(* IEC 61131-3 sources: TIA2AX/tests/test_projects/expected/HW_DiscoverGroups/PLC_2, 6 files *)

(* ---- HwInputs.st ---- *)
TYPE
	HwInputs : STRUCT
		PLC_2_10A_1 AT %B7 : WORD;
		PLC_2_10A_2 AT %B9 : WORD;
		PLC_2_10A_3 AT %B11 : WORD;
		PLC_2_10A_4 AT %B13 : WORD;
		PLC_2_10A_5 AT %B15 : WORD;
		PLC_2_10A_6 AT %B17 : WORD;
		_10A_16_10A_2 AT %B19 : BYTE;
		_10A_16_10A_3 AT %B20 : BYTE;
		_10A_16_10A_4 AT %B21 : BYTE;
		_10A_16_10A_5 AT %B22 : BYTE;
		_10A_16_10A_6 AT %B23 : BYTE;
		_10A_20_10A_2 AT %B24 : BYTE;
		_10A_20_10A_3 AT %B25 : BYTE;
		_10A_20_10A_4 AT %B26 : BYTE;
		_10A_20_10A_5 AT %B27 : BYTE;
		_10A_20_10A_6 AT %B28 : BYTE;
		_10A_12_10A_2 AT %B2 : BYTE;
		_10A_12_10A_3 AT %B3 : BYTE;
		_10A_12_10A_4 AT %B4 : BYTE;
		_10A_12_10A_5 AT %B5 : BYTE;
		_10A_12_10A_6 AT %B6 : BYTE;
	END_STRUCT;
END_TYPE

(* ---- HwOutputs.st ---- *)
TYPE
	HwOutputs : STRUCT
		PLC_2_10A_7 AT %B7 : WORD;
		PLC_2_10A_8 AT %B9 : WORD;
		PLC_2_10A_9 AT %B11 : WORD;
		PLC_2_10A_10 AT %B13 : WORD;
		PLC_2_10A_11 AT %B15 : WORD;
		PLC_2_10A_12 AT %B17 : WORD;
		_10A_16_10A_7 AT %B19 : BYTE;
		_10A_16_10A_8 AT %B20 : BYTE;
		_10A_16_10A_9 AT %B21 : BYTE;
		_10A_16_10A_10 AT %B22 : BYTE;
		_10A_16_10A_11 AT %B23 : BYTE;
		_10A_20_10A_7 AT %B24 : BYTE;
		_10A_20_10A_8 AT %B25 : BYTE;
		_10A_20_10A_9 AT %B26 : BYTE;
		_10A_20_10A_10 AT %B27 : BYTE;
		_10A_20_10A_11 AT %B28 : BYTE;
		_10A_12_10A_7 AT %B2 : BYTE;
		_10A_12_10A_8 AT %B3 : BYTE;
		_10A_12_10A_9 AT %B4 : BYTE;
		_10A_12_10A_10 AT %B5 : BYTE;
		_10A_12_10A_11 AT %B6 : BYTE;
	END_STRUCT;
END_TYPE

(* ---- PlcInputs.st ---- *)
TYPE
	PlcInputs : STRUCT
		PLC_2_10A_1 : WORD;
		PLC_2_10A_2 : WORD;
		PLC_2_10A_3 : WORD;
		PLC_2_10A_4 : WORD;
		PLC_2_10A_5 : WORD;
		PLC_2_10A_6 : WORD;
		_10A_16_10A_2 : BYTE;
		_10A_16_10A_3 : BYTE;
		_10A_16_10A_4 : BYTE;
		_10A_16_10A_5 : BYTE;
		_10A_16_10A_6 : BYTE;
		_10A_20_10A_2 : BYTE;
		_10A_20_10A_3 : BYTE;
		_10A_20_10A_4 : BYTE;
		_10A_20_10A_5 : BYTE;
		_10A_20_10A_6 : BYTE;
		_10A_12_10A_2 : BYTE;
		_10A_12_10A_3 : BYTE;
		_10A_12_10A_4 : BYTE;
		_10A_12_10A_5 : BYTE;
		_10A_12_10A_6 : BYTE;
	END_STRUCT;
END_TYPE

(* ---- PlcOutputs.st ---- *)
TYPE
	PlcOutputs : STRUCT
		PLC_2_10A_7 : WORD;
		PLC_2_10A_8 : WORD;
		PLC_2_10A_9 : WORD;
		PLC_2_10A_10 : WORD;
		PLC_2_10A_11 : WORD;
		PLC_2_10A_12 : WORD;
		_10A_16_10A_7 : BYTE;
		_10A_16_10A_8 : BYTE;
		_10A_16_10A_9 : BYTE;
		_10A_16_10A_10 : BYTE;
		_10A_16_10A_11 : BYTE;
		_10A_20_10A_7 : BYTE;
		_10A_20_10A_8 : BYTE;
		_10A_20_10A_9 : BYTE;
		_10A_20_10A_10 : BYTE;
		_10A_20_10A_11 : BYTE;
		_10A_12_10A_7 : BYTE;
		_10A_12_10A_8 : BYTE;
		_10A_12_10A_9 : BYTE;
		_10A_12_10A_10 : BYTE;
		_10A_12_10A_11 : BYTE;
	END_STRUCT;
END_TYPE

(* ---- CopyInputs.st ---- *)
FUNCTION CopyInputs
	VAR_EXTERNAL
		HwInputs : HwInputs;
		PlcInputs : PlcInputs;
	END_VAR
	PlcInputs.PLC_2_10A_1 := HwInputs.PLC_2_10A_1;
	PlcInputs.PLC_2_10A_2 := HwInputs.PLC_2_10A_2;
	PlcInputs.PLC_2_10A_3 := HwInputs.PLC_2_10A_3;
	PlcInputs.PLC_2_10A_4 := HwInputs.PLC_2_10A_4;
	PlcInputs.PLC_2_10A_5 := HwInputs.PLC_2_10A_5;
	PlcInputs.PLC_2_10A_6 := HwInputs.PLC_2_10A_6;
	PlcInputs._10A_16_10A_2 := HwInputs._10A_16_10A_2;
	PlcInputs._10A_16_10A_3 := HwInputs._10A_16_10A_3;
	PlcInputs._10A_16_10A_4 := HwInputs._10A_16_10A_4;
	PlcInputs._10A_16_10A_5 := HwInputs._10A_16_10A_5;
	PlcInputs._10A_16_10A_6 := HwInputs._10A_16_10A_6;
	PlcInputs._10A_20_10A_2 := HwInputs._10A_20_10A_2;
	PlcInputs._10A_20_10A_3 := HwInputs._10A_20_10A_3;
	PlcInputs._10A_20_10A_4 := HwInputs._10A_20_10A_4;
	PlcInputs._10A_20_10A_5 := HwInputs._10A_20_10A_5;
	PlcInputs._10A_20_10A_6 := HwInputs._10A_20_10A_6;
	PlcInputs._10A_12_10A_2 := HwInputs._10A_12_10A_2;
	PlcInputs._10A_12_10A_3 := HwInputs._10A_12_10A_3;
	PlcInputs._10A_12_10A_4 := HwInputs._10A_12_10A_4;
	PlcInputs._10A_12_10A_5 := HwInputs._10A_12_10A_5;
	PlcInputs._10A_12_10A_6 := HwInputs._10A_12_10A_6;
END_FUNCTION

(* ---- CopyOutputs.st ---- *)
FUNCTION CopyOutputs
	VAR_EXTERNAL
		HwOutputs : HwOutputs;
		PlcOutputs : PlcOutputs;
	END_VAR
	HwOutputs.PLC_2_10A_7 := PlcOutputs.PLC_2_10A_7;
	HwOutputs.PLC_2_10A_8 := PlcOutputs.PLC_2_10A_8;
	HwOutputs.PLC_2_10A_9 := PlcOutputs.PLC_2_10A_9;
	HwOutputs.PLC_2_10A_10 := PlcOutputs.PLC_2_10A_10;
	HwOutputs.PLC_2_10A_11 := PlcOutputs.PLC_2_10A_11;
	HwOutputs.PLC_2_10A_12 := PlcOutputs.PLC_2_10A_12;
	HwOutputs._10A_16_10A_7 := PlcOutputs._10A_16_10A_7;
	HwOutputs._10A_16_10A_8 := PlcOutputs._10A_16_10A_8;
	HwOutputs._10A_16_10A_9 := PlcOutputs._10A_16_10A_9;
	HwOutputs._10A_16_10A_10 := PlcOutputs._10A_16_10A_10;
	HwOutputs._10A_16_10A_11 := PlcOutputs._10A_16_10A_11;
	HwOutputs._10A_20_10A_7 := PlcOutputs._10A_20_10A_7;
	HwOutputs._10A_20_10A_8 := PlcOutputs._10A_20_10A_8;
	HwOutputs._10A_20_10A_9 := PlcOutputs._10A_20_10A_9;
	HwOutputs._10A_20_10A_10 := PlcOutputs._10A_20_10A_10;
	HwOutputs._10A_20_10A_11 := PlcOutputs._10A_20_10A_11;
	HwOutputs._10A_12_10A_7 := PlcOutputs._10A_12_10A_7;
	HwOutputs._10A_12_10A_8 := PlcOutputs._10A_12_10A_8;
	HwOutputs._10A_12_10A_9 := PlcOutputs._10A_12_10A_9;
	HwOutputs._10A_12_10A_10 := PlcOutputs._10A_12_10A_10;
	HwOutputs._10A_12_10A_11 := PlcOutputs._10A_12_10A_11;
END_FUNCTION
